FUNCTION_BLOCK invert_output (* Basic Function Block Type *)
  (* Standard: 61499-2 *)
  (* Version 0.0, 12/30/2019, prana, nxtControl GmbH, Template *)
  PACKAGE Main;
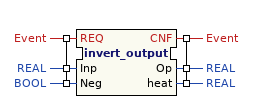
  EVENT_INPUT
    REQ WITH Inp, Neg; (* Normal Execution Request *)
  END_EVENT
  EVENT_OUTPUT
    CNF WITH Op, heat; (* Execution Confirmation *)
  END_EVENT
  VAR_INPUT
    Inp : REAL; (* Input event qualifier *)
    Neg : BOOL;
  END_VAR
  VAR_OUTPUT
    Op : REAL; (* Output event qualifier *)
    heat : REAL;
  END_VAR
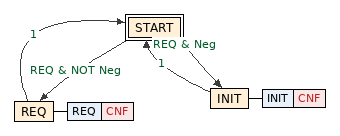
  EC_STATES
    START; (* Initial State *)
    INIT : INIT -> CNF; (* Initialization *)
    REQ : REQ -> CNF; (* Normal execution *)
  END_STATES
  EC_TRANSITIONS
    START TO INIT := REQ & Neg;
    INIT TO START := 1;
    START TO REQ := REQ & NOT Neg;
    REQ TO START := 1;
  END_TRANSITIONS
  ALGORITHM INIT IN ST: (* Initialization algorithm *)
Op := -Inp;
heat := 0;
  END_ALGORITHM
  ALGORITHM REQ IN ST: (* Normally executed algorithm *)
Op :=  Inp;
heat := 1;
  END_ALGORITHM
END_FUNCTION_BLOCK
